(* IEC 61131-3 sources: Elmo_Master/Lasal_PRG/MotionTCPDemo/Network/UDPComNet, 1 file *)

(* ---- ONE_UDPComNet_Table.st ---- *)
#define OBJECTS_CONFIG

//Define part of class _UDPTransceiver
#define UDP_MAX_SOCKETS               6                             // Max number of socket

#define UDP_CLT_SEND_OK               0                             // Send ok
#define UDP_CLT_INVALID_HANDLE        -1                            // Invalid handle
#define UDP_CLT_NOT_OPEN              -2                            // Socket is not open
#define UDP_CLT_SEND_FAILED           -3                            // Send failed
#define UDP_CLT_SEND_BUFFER_FULL      -4                            // Send buffer is full
#define UDP_CLT_DATA_TO_BIG           -5                            // Data to big
#define UDP_CLT_INVALID_DATA          -6

#define UDP_MAXIMUM_SEGMENT_SIZE      1452                          //

#define MAX_MSG_CYC_SEND                5
#define MAX_MSG_CYC_RECV                5

#define UDP_CLT_INFO_ADDED          0
#define UDP_CLT_INFO_BOUND          1
#define UDP_CLT_INFO_CLOSED         2
#include <.\lsl_st_mt.h>
//Define part of class UDPTransmission
#define IP_ADDR_MIN_LEN         7
#define IP_ADDR_MAX_LEN         15

FUNCTION GLOBAL TAB ONE_UDPComNet
-1$UINT, 0$UINT,
0$UINT, 0$UINT,

8$UDINT,
TO_UDINT(3808005437), "_UDPTransceiver", 1$UINT, 2$UINT, 1$UINT,
TO_UDINT(3441197119), "_UDPTransceiverInterface", 1$UINT, 3$UINT, 0$UINT,
TO_UDINT(794617671), "CriticalSection", 0$UINT, 4$UINT, 2$UINT,
TO_UDINT(2225119864), "MerkerEx", 1$UINT, 22$UINT, 1$UINT,
TO_UDINT(1850111279), "String", 1$UINT, 11$UINT, 1$UINT,
TO_UDINT(2898603620), "StringInternal", 1$UINT, 86$UINT, 0$UINT,
TO_UDINT(2855436325), "UDPTransmission", 0$UINT, 0$UINT, 1$UINT,
TO_UDINT(3232495061), "VirtualBaseInit", 1$UINT, 3$UINT, 0$UINT,

_NO_ATTR, TO_UDINT(3679869483), "_UDPTRANSCEIVER1",

1$UINT, TO_UDINT(152563782), "UDPTRANSMISSION1\_BASE\CRITICALSECTION_UDP",
1$UINT, TO_UDINT(936750719), "_UDPTRANSCEIVER1\CRITICALSECTION_UDP",

1$UINT, TO_UDINT(3025948), "STRING1\MERKEREX0",

_NO_ATTR, TO_UDINT(677614747), "STRING1",

_NO_ATTR, TO_UDINT(3362916720), "UDPTRANSMISSION1",

//Internal connections
0$UDINT,
3$UDINT,
TO_UDINT(0), "CriticalSection_UDP", TO_UDINT(2),
TO_UDINT(4), "MerkerEx0", TO_UDINT(3),
TO_UDINT(5), "CriticalSection_UDP", TO_UDINT(1),
0$UDINT,
3$UDINT,
TO_UDINT(4), "DataBuffer", TO_UDINT(3), "m_udLength",
TO_UDINT(5), "_UDPTransceiver", TO_UDINT(0), "sControl",
TO_UDINT(5), "IPAddr", TO_UDINT(4), "Data",

//Initialization values
0$UDINT,
5$UDINT,
TO_UDINT(0), "cSizeOfTXBuffer", TO_UDINT(100 kb),//|UDPComNet._UDPTransceiver1.cSizeOfTXBuffer;
TO_UDINT(0), "cSizeOfRXBuffer", TO_UDINT(100 kb),//|UDPComNet._UDPTransceiver1.cSizeOfRXBuffer;
TO_UDINT(3), "ThreadSafe", TO_UDINT(0),//|UDPComNet.String1\MerkerEx0.ThreadSafe;
TO_UDINT(4), "SingleRealloc", TO_UDINT(1),//|UDPComNet.String1.SingleRealloc;
TO_UDINT(5), "Port", TO_UDINT(8877),//|UDPComNet.UDPTransmission1.Port;

//Symbolic initialization values
0$UDINT,
0$UDINT,

//Initialization of string values
0$UDINT,
1$UDINT,
TO_UDINT(4), "", 0$UINT, TO_UINT(OFF(L1)-OFF(L0)), L0:"192.168.111.101",L1://|UDPComNet.String1.Data;

//Configuration of tasks (RealTime, Cyclic, Background)
0$UDINT,
0$UDINT,

0$UDINT,
2$UDINT,
TO_UDINT(0), (1)$UDINT, 4194303$DINT, 	//_UDPTRANSCEIVER1
TO_UDINT(5), (10)$UDINT, 4194303$DINT, 	//UDPTRANSMISSION1

0$UDINT,
0$UDINT,

//External connections
0$UDINT,
0$UDINT,

//Magic internal connections
0$UDINT,
0$UDINT,

//Configuration of timeslots of tasks (RealTime, Cyclic)
#ifdef __LSLLDR_TIMESLOTS__
0$UDINT,
0$UDINT,

0$UDINT,
0$UDINT,

#endif //__LSLLDR_TIMESLOTS__

//MultiMaster connections
#ifdef __LSLLDR_MULTIMASTER__
0$UDINT,
0$UDINT,
#endif //__LSLLDR_MULTIMASTER__

//Configuration for task ID (RealTime, CyclicTime)
#ifdef __LSLLDR_TASKID__
"\\\\TASKS2  "
0$UDINT,
0$UDINT,

0$UDINT,
2$UDINT,
(0)$UDINT, 	//_UDPTRANSCEIVER1
(0)$UDINT, 	//UDPTRANSMISSION1

0$UDINT,
0$UDINT,

#endif //__LSLLDR_TASKID__

END_FUNCTION
